(* IEC 61131-3 sources: kns-port-domestic/upstream/kns-pump-station/src/DUTs/Sim, 9 files *)

(* ---- E_SimAiFault.dut.st ---- *)
// Назначение: инъекция отказа аналогового датчика 4–20 мА в модели (NAMUR NE 43): обрыв,
//             токи отказа и выхода из диапазона, замерзание, принудительный ток.
// Автор:      kr0nsch
// Версия:     0.1.0
// Документ:   docs/DESIGN.md, раздел 3.3; docs/06_PMI.md, раздел 5.4
{attribute 'qualified_only'}
{attribute 'strict'}
TYPE E_SimAiFault :
(
    None := 0,          // нет инъекции: ток по измеренному значению
    WireBreak := 1,     // обрыв линии: 0 мА
    FailLow := 2,       // отказ снизу: SIM_MA_FAIL_LOW (3,0 мА)
    FailHigh := 3,      // отказ сверху: SIM_MA_FAIL_HIGH (22 мА)
    UnderRange := 4,    // ниже диапазона: SIM_MA_UNDER_RANGE (3,7 мА)
    OverRange := 5,     // выше диапазона: SIM_MA_OVER_RANGE (20,8 мА)
    Freeze := 6,        // замерзание: последнее значение тока
    Forced := 7         // принудительный ток arAiForced_mA
) INT;
END_TYPE

(* ---- E_SimFloatStuck.dut.st ---- *)
// Назначение: инъекция залипания поплавкового выключателя в модели.
// Автор:      kr0nsch
// Версия:     0.1.0
// Документ:   docs/DESIGN.md, раздел 3.3; docs/06_PMI.md, раздел 5.4
{attribute 'qualified_only'}
{attribute 'strict'}
TYPE E_SimFloatStuck :
(
    None := 0,          // нет инъекции: контакт по уровню
    StuckNormal := 1,   // контакт не срабатывает (НЗ остаётся замкнутым)
    StuckTripped := 2   // сработал и не возвращается; то же — обрыв цепи НЗ-контакта
) INT;
END_TYPE

(* ---- ST_FaultInjection.dut.st ---- *)
// Назначение: инъекции отказов модели (GVL_Sim.stFaultInj). Пишут HMI (экран «Имитация») и
//             сценарии ПМИ; действуют только при GVL_Sim.xSimulation. Индекс насоса 1…3 = Н1…Н3,
//             индекс датчика — SIM_AI_*. Имена полей использует таблица 06 §5.4 и экран 08.
// Автор:      kr0nsch
// Версия:     0.1.0
// Документ:   docs/DESIGN.md, раздел 3.3; docs/06_PMI.md, раздел 5.4
{attribute 'qualified_only'}
TYPE ST_FaultInjection :
STRUCT
    // авария ПЧ: реле FLT, бит STW.2, код SIM_VFD_FCODE_EXT; снимается сбросом ПЧ после снятия инъекции
    axVfdFault      : ARRAY[1..GVL_Const.STN_PUMP_COUNT] OF BOOL;
    // реле «Работа» не замыкается (ПЧ работает) → FailToStart / FeedbackLost
    axNoFeedback    : ARRAY[1..GVL_Const.STN_PUMP_COUNT] OF BOOL;
    // реле «Работа» залипло в TRUE → FailToStop / UncommandedRun
    axFeedbackStuck : ARRAY[1..GVL_Const.STN_PUMP_COUNT] OF BOOL;
    axAirLock       : ARRAY[1..GVL_Const.STN_PUMP_COUNT] OF BOOL;  // сухой ход насоса: подача 0, ток мал → недогрузка
    axClog          : ARRAY[1..GVL_Const.STN_PUMP_COUNT] OF BOOL;  // засор: подача −60 %, ток ×1,3 к току без засора
    axOverheat      : ARRAY[1..GVL_Const.STN_PUMP_COUNT] OF BOOL;  // TS1n2 размыкается и разрывает цепь аварии ПЧ
    axLeak          : ARRAY[1..GVL_Const.STN_PUMP_COUNT] OF BOOL;  // MS1n3
    // нет ответа ПЧ: регистры замирают, xMbOk = FALSE; через SIM_VFD_WATCHDOG — 50 Гц (04 §12);
    // все три — потеря линии RS485-1
    axVfdCommLoss   : ARRAY[1..GVL_Const.STN_PUMP_COUNT] OF BOOL;
    axLocal         : ARRAY[1..GVL_Const.STN_PUMP_COUNT] OF BOOL;  // переключатель HS1n4 в «Местное»
    axLocalRun      : ARRAY[1..GVL_Const.STN_PUMP_COUNT] OF BOOL;  // пуск с местного поста (в «Местном»)
    // индексы SIM_AI_*: LT101, PT201, FT202, AT401, AT402
    aeAiFault       : ARRAY[1..GVL_Const.SIM_AI_COUNT] OF E_SimAiFault;
    arAiForced_mA   : ARRAY[1..GVL_Const.SIM_AI_COUNT] OF REAL;  // ток при Forced
    eLs102Stuck     : E_SimFloatStuck;
    eLs103Stuck     : E_SimFloatStuck;
    xPowerLoss      : BOOL;                 // нет напряжения на вводе: ES301 = 0, ПЧ обесточены, ИБП на батареях
    xUpsFault       : BOOL;                 // YS303
    xTempCommLoss   : BOOL;                 // TT403 (RS485-2) не отвечает
    xFanFault       : BOOL;                 // V1_FLT
    xFanNoFeedback  : BOOL;                 // V1_RFB не приходит при работающем вентиляторе (04 §20, вопрос 10)
    xValveChamberFlood : BOOL;              // LS203
    xFire           : BOOL;                 // YS405
    // концентрации газов вместо фоновых из stSimCfg; < 0 — фон (по умолчанию и после xClearFaults)
    rH2S_mgm3       : REAL := -1.0;
    rCh4_pctLel     : REAL := -1.0;
END_STRUCT
END_TYPE

(* ---- ST_PlantIo.dut.st ---- *)
// Назначение: все сигналы модели для входов GVL_IO: входы модулей AI/DI, регистры чтения ПЧ и
//             TT403, состояние обмена со слейвами Modbus. Поля называются так же, как переменные
//             GVL_IO (вывод iolistgen по docs/03_io_list.csv): PRG_PlantModel копирует поле в
//             одноимённую переменную. Модель пишет только входы GVL_IO (ARCHITECTURE, раздел 4).
// Автор:      kr0nsch
// Версия:     0.1.0
// Документ:   docs/DESIGN.md, разделы 3.3, 11.1; docs/03_io_list.md
{attribute 'qualified_only'}
TYPE ST_PlantIo :
STRUCT
    // --- входы AI, мА ---
    rLT101_mA : REAL;               // A1.1 уровень, 0…5 м
    rPT201_mA : REAL;               // A1.2 давление в коллекторе, 0…10 бар
    rFT202_mA : REAL;               // A1.3 расход, 0…500 м³/ч
    rAT401_mA : REAL;               // A1.4 H2S, 0…40 мг/м³
    rAT402_mA : REAL;               // A1.5 CH4, 0…100 % НКПР
    // --- входы DI шкафа и павильона ---
    xLS102 : BOOL;                  // поплавок «аварийно высокий», НЗ: TRUE — норма
    xLS103 : BOOL;                  // поплавок «сухой ход», НЗ: TRUE — норма
    xLS203 : BOOL;                  // затопление камеры задвижек
    xES301 : BOOL;                  // напряжение на вводе в норме
    xYS302 : BOOL;                  // ИБП: работа от батарей
    xYS303 : BOOL;                  // ИБП: неисправность
    xZS404 : BOOL;                  // дверь павильона открыта
    xYS405 : BOOL;                  // пожар
    xHS501 : BOOL;                  // кнопка «Сброс аварий»
    xHS502 : BOOL;                  // кнопка «Отключить звук»
    xV1_RFB : BOOL;                 // В1: блок-контакт пускателя
    xV1_FLT : BOOL;                 // В1: автомат защиты двигателя
    // --- входы DI насосов ---
    xP101_RFB : BOOL;               // Н1: реле ПЧ «Работа»
    xP101_FLT : BOOL;               // Н1: реле ПЧ «Авария»
    xHS114 : BOOL;                  // Н1: «Местное»
    xTS112 : BOOL;                  // Н1: термовыключатели, НЗ: TRUE — норма
    xMS113 : BOOL;                  // Н1: протечка в камеру статора
    xP102_RFB : BOOL;
    xP102_FLT : BOOL;
    xHS124 : BOOL;
    xTS122 : BOOL;
    xMS123 : BOOL;
    xP103_RFB : BOOL;
    xP103_FLT : BOOL;
    xHS134 : BOOL;
    xTS132 : BOOL;
    xMS133 : BOOL;
    // --- регистры чтения ПЧ (RS485-1, FC3 100…103) ---
    wP101_STW : WORD;               // слово состояния
    uiP101_FACT : UINT;             // фактическая частота, 0,01 Гц
    uiIT111 : UINT;                 // ток двигателя, 0,1 А
    uiP101_FCODE : UINT;            // код последней аварии
    wP102_STW : WORD;
    uiP102_FACT : UINT;
    uiIT121 : UINT;
    uiP102_FCODE : UINT;
    wP103_STW : WORD;
    uiP103_FACT : UINT;
    uiIT131 : UINT;
    uiP103_FCODE : UINT;
    // --- RS485-2: температура павильона ---
    rTT403 : REAL;                  // °C
    // --- состояние обмена со слейвами ---
    xMbOk_RS485_1_S1 : BOOL;
    xMbOk_RS485_1_S2 : BOOL;
    xMbOk_RS485_1_S3 : BOOL;
    xMbOk_RS485_2_S10 : BOOL;
END_STRUCT
END_TYPE

(* ---- ST_PumpModelCfg.dut.st ---- *)
// Назначение: характеристика насоса и сети для модели (законы подобия, рабочая точка, ток
//             двигателя). Значения по умолчанию — условные, подобраны под подачи документов
//             (DESIGN 11.3; сверяет эталон tools_project/plant_reference.py).
// Автор:      kr0nsch
// Версия:     0.1.0
// Документ:   docs/DESIGN.md, разделы 3.3, 11.2, 11.3
{attribute 'qualified_only'}
TYPE ST_PumpModelCfg :
STRUCT
    rH0_m      : REAL := 34.5;      // напор при нулевой подаче на 50 Гц
    rK_mh2     : REAL := 6.06E-4;   // крутизна характеристики, м/(м³/ч)²
    rHgeo_m    : REAL := 12.0;      // геометрический напор от дна резервуара
    rR_mh2     : REAL := 4.60E-4;   // сопротивление трубопровода, м/(м³/ч)²
    rEta       : REAL := 0.62;      // КПД агрегата
    rPnom_kW   : REAL := 15.0;
    rInom_A    : REAL := 28.0;
    rImagShare : REAL := 0.30;      // доля намагничивающего тока
    rLossShare : REAL := 0.12;      // потери без подачи, доля Pnom
END_STRUCT
END_TYPE

(* ---- ST_SimCfg.dut.st ---- *)
// Назначение: параметры модели и ускорение контура (GVL_Sim.stSimCfg). Значения по умолчанию —
//             условные (DESIGN 11.3), согласованы с 04 и 06.
// Автор:      kr0nsch
// Версия:     0.1.0
// Документ:   docs/DESIGN.md, разделы 3.3, 11.3
{attribute 'qualified_only'}
TYPE ST_SimCfg :
STRUCT
    rTimeScale        : REAL := 1.0;        // 1…SIM_TIME_SCALE_MAX: ускорение всего контура (ARCHITECTURE, раздел 11)
    rTankArea_m2      : REAL := 12.0;
    rLevelOverflow_m  : REAL := 4.60;
    rLevelInit_m      : REAL := 1.20;
    rInflowAvg_m3h    : REAL := 70.0;
    arDailyProfile    : ARRAY[0..GVL_Const.SIM_PROFILE_POINTS - 1] OF REAL := [0.55, 0.45, 0.40, 0.38, 0.40, 0.55,
                            0.92, 1.35, 1.60, 1.50, 1.30, 1.15, 1.10, 1.05, 1.00, 1.00, 1.00, 1.15, 1.35, 1.50,
                            1.45, 1.20, 0.95, 0.70];
    udiSeed           : UDINT := 20261016;  // генератор ливней (одинаковый seed — одинаковые ливни)
    uiStormsPerDayMax : UINT := 2;          // не больше SIM_STORMS_MAX
    rStormPeakMin_m3h : REAL := 100.0;
    rStormPeakMax_m3h : REAL := 250.0;
    tStormMin         : TIME := T#20M;
    tStormMax         : TIME := T#90M;
    rStartTimeOfDay_h : REAL := 0.0;        // время суток модели при старте; демонстрация задаёт его командой
    stPump            : ST_PumpModelCfg;
    tVfdAccel         : TIME := T#10S;      // разгон ПЧ 0 → 50 Гц
    tVfdBoot          : TIME := T#5S;       // готовность ПЧ после подачи питания
    rH2SBase_mgm3     : REAL := 0.6;        // фон газов и температура павильона (условно)
    rCh4Base_pctLel   : REAL := 1.5;
    rAirTemp_C        : REAL := 18.0;
END_STRUCT
END_TYPE

(* ---- ST_SimCmd.dut.st ---- *)
// Назначение: команды модели (GVL_Sim.stSimCmd). Импульсы сбрасывает модель (FB_PlantModel)
//             после выполнения; xInflowOverride и xDoorOpen — уровни.
// Автор:      kr0nsch
// Версия:     0.1.0
// Документ:   docs/DESIGN.md, раздел 3.3; docs/06_PMI.md, раздел 5.4
{attribute 'qualified_only'}
TYPE ST_SimCmd :
STRUCT
    xResetPlant      : BOOL;        // импульс: уровень := stSimCfg.rLevelInit_m, перелив 0, ливни сняты, ПЧ готовы
    xClearFaults     : BOOL;        // импульс: обнулить stFaultInj (ускорение и приток не меняются)
    xSetLevel        : BOOL;        // импульс: уровень := rSetLevel_m
    rSetLevel_m      : REAL;
    xInflowOverride  : BOOL;        // уровень: приток := rInflowOverride_m3h (без профиля и ливней)
    rInflowOverride_m3h : REAL;
    xStormNow        : BOOL;        // импульс: ливень сейчас (при xInflowOverride = FALSE)
    rStormPeak_m3h   : REAL;
    tStormDuration   : TIME;
    xSetTimeOfDay    : BOOL;        // импульс: время суток модели := rTimeOfDay_h
    rTimeOfDay_h     : REAL;
    xPressReset      : BOOL;        // импульс: нажать HS501 на SIM_BUTTON_PULSE
    xPressSilence    : BOOL;        // импульс: нажать HS502
    xDoorOpen        : BOOL;        // уровень: дверь павильона открыта (ZS404)
END_STRUCT
END_TYPE

(* ---- ST_SimSts.dut.st ---- *)
// Назначение: состояние модели (GVL_Sim.stSimSts, только чтение): истинный уровень, потоки,
//             частоты и токи насосов, время суток, ливни, перелив, счётчик изменений инъекций.
// Автор:      kr0nsch
// Версия:     0.1.0
// Документ:   docs/DESIGN.md, раздел 3.3
{attribute 'qualified_only'}
TYPE ST_SimSts :
STRUCT
    rLevel_m         : REAL;        // истинный уровень
    rInflow_m3h      : REAL;
    rOutflow_m3h     : REAL;
    arPumpFlow_m3h   : ARRAY[1..GVL_Const.STN_PUMP_COUNT] OF REAL;
    rHead_m          : REAL;
    arFreq_Hz        : ARRAY[1..GVL_Const.STN_PUMP_COUNT] OF REAL;
    arCurrent_A      : ARRAY[1..GVL_Const.STN_PUMP_COUNT] OF REAL;
    rTimeOfDay_h     : REAL;
    udiDay           : UDINT;
    xStormActive     : BOOL;
    rStormInflow_m3h : REAL;
    udiOverflow_s    : UDINT;       // время перелива (время контура)
    rTimeScaleAct    : REAL;
    lrSimTime_s      : LREAL;
    xRunning         : BOOL;        // модель работает
    udiFaultSeq      : UDINT;       // +1 при каждом изменении stFaultInj; по нему PRG_Station пишет событие 101021
END_STRUCT
END_TYPE

(* ---- ST_StormEvent.dut.st ---- *)
// Назначение: ливень генератора модели: начало в сутках, длительность, пик притока
//             (форма — трапеция: рост 15 %, полка 50 %, спад 35 % длительности).
// Автор:      kr0nsch
// Версия:     0.1.0
// Документ:   docs/DESIGN.md, разделы 3.3, 11.2
{attribute 'qualified_only'}
TYPE ST_StormEvent :
STRUCT
    rStart_h  : REAL;               // начало, ч от полуночи суток
    tDuration : TIME;
    rPeak_m3h : REAL;
END_STRUCT
END_TYPE
